FUNCTION_BLOCK T_Test1 EXTENDS T_UnitTestBase IMPLEMENTS I_UnitTest
VAR
	Value : INT := 7;
END_VAR

{attribute 'analysis' := '-33'} // inhibit unused variable warning
METHOD  RunTest
VAR_INST
	OnTimer : T_OnTimer(PresetTime := 1.5);
END_VAR
CASE State OF
    0:
        OnTimer.Reset();
        Value := 5;
        F_Inc(State);
    1:
        AssertEquals_INT(Expected := 7, Actual := Value, Message := 'Value');
        F_Inc(State);

    2:
        IF OnTimer.Run() THEN
            _Completed := TRUE;
        END_IF

END_CASE
END_METHOD

END_FUNCTION_BLOCK

(* stored: Version 1.1.0.1, ProductVersion 3.1.4024.15
   POU T_Test1: Id {38fce957-6a84-4940-8b00-735d0a8d36e5}, SpecialFunc None
   Method RunTest: Id {4703f096-77af-4272-9877-be9134bb7616} *)
